(* Logix 5000 project; controller TFF vendor 1 type 14 code 107 rev 33.11; software revision 33.04; part 36 of 38 *)
(* tags used below, declared in another part *)
   Address : DINT;   // Temp Address
   AlarmInhibit_Timer : TIMER;
   Index : DINT;   // Index
   NewSystem : DINT;
   TIME : DINT[2];
   AI201B : ALIAS FOR AnalogPoint[0];
   AI201BAlarm : ALIAS FOR AlarmAnalog[0];
   AlarmAnalog_Storage : AlarmAnalog[6,50];
   AlarmDeviation : AlarmDeviation[20];   // Control Loop Deviation Alarm Array
   AlarmDeviation_Storage : AlarmDeviation[6,20];
   AnalogOutput_Storage : AnalogOutput[6,25];
   AnalogPoint_Storage : AnalogInput[6,50];
   CCPSystem : CCPSystem;   // CCP System Data
   CCPSystem_Storage : CCPSystem_Storage[6];
   ControlLoop : ControlLoop[20];   // Control Loop Array
   ControlLoop_Storage : ControlLoop[6,20];
   DigitalPoint_Storage : DigitalPoint[6,150];
   Drive : Drive[11];   // Drives Array
   Drive_Storage : Drive[6,11];
   FlowPath : FlowPath[64];   // Flow Path Array
   FlowPath_Storage : FlowPath[6,64];
   Gateway : Gateway;   // Gateway Control
   GWModbus : IO_Station;   // Status of Gateway Modbus
   Options : Options;   // Options List
   Phase0 : ALIAS FOR Phase[0];   // Phase 0
   Phase0_Totalizer_Feed : ALIAS FOR PhaseTotalizer[0];   // Phase 0 Total Feed
   PhaseTotalizer : PhaseTotalizer[18];   // Phase Totalizers Array
   PhaseTotalizer_Storage : PhaseTotalizer[6,18];
   PipeAnimation : PipeAnimation;   // HMI Pipe Animation Array
   PipeStatValueHMI : INT[224];   // Pipe Animation Value For HMI
   PISL601 : ALIAS FOR DigitalPoint[0];
   Rack_ACT350_WI101_200L : IO_Station;   // Status of ACT350 200L
   Rack_ACT350_WI101_500L : IO_Station;   // Status of ACT350 500L
   Rack_Murr_Node0_Smart : IO_Station;   // Status of Node 0 Smart
   Rack_Murr_Node1_TFF20 : IO_Station;   // Status of Node 1 TFF20
   Rack_Murr_Node1_TFF40 : IO_Station;   // Status of Node 1 TFF40
   Rack_Murr_Node1_TFF80 : IO_Station;   // Status of Node 1 TFF80
   SIC001 : ALIAS FOR Drive[1];
   SIC001_AO : ALIAS FOR AnalogOutput[0];
   SIC002 : ALIAS FOR Drive[2];
   ThisSystem : SystemType;
   Valve_Storage : Valve[6,100];
   WI101 : ALIAS FOR AnalogPoint[15];
   XV001 : ALIAS FOR Valve[0];
(* Process, continued *)

ROUTINE PipeAnimationHMI   (* ladder *)
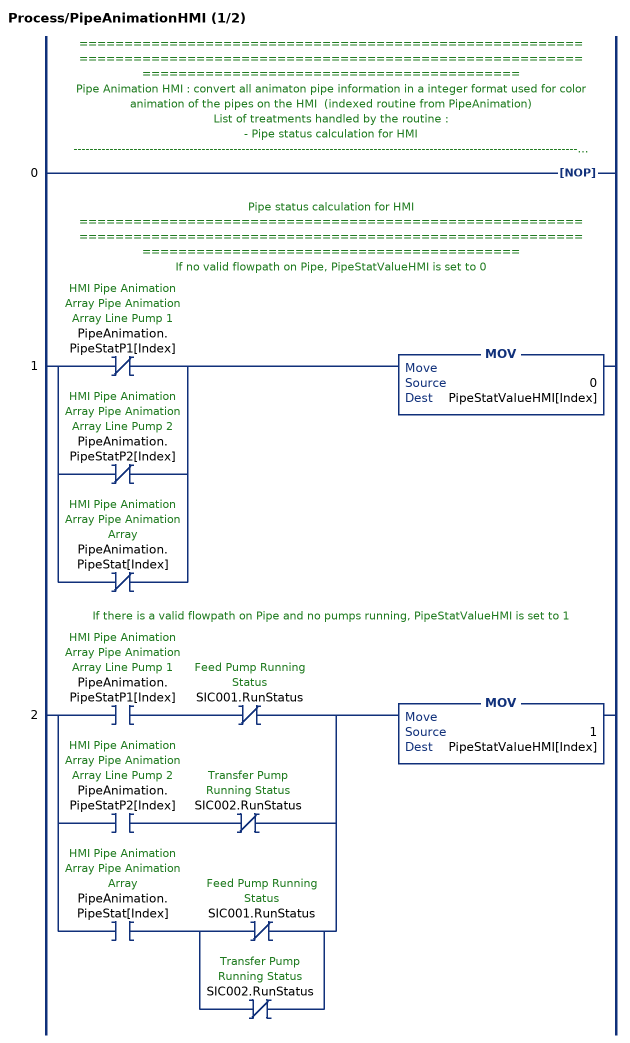
   // ==========================================================================================================================================================
   //                          Pipe Animation HMI : convert all animaton pipe information in a integer format used for color animation of the pipes on the HMI  (indexed routine from PipeAnimation)
   //                                                     List of treatments handled by the routine :
   //                                                          - Pipe status calculation for HMI
   //                                                     -----------------------------------------------------------------------------------------------------------------------------------------------------
   //                                                     History
   // 		2019-DEC-24 - Merck - Q. Spindler - Initial version for Candidate Release 1.00.00.00.a
   // ========================================================================================================================================================
   0: NOP();
   // Pipe status calculation for HMI
   // ==========================================================================================================================================================
   // If no valid flowpath on Pipe, PipeStatValueHMI is set to 0
   1: [XIO(PipeAnimation.PipeStatP1[Index]) ,XIO(PipeAnimation.PipeStatP2[Index]) ,XIO(PipeAnimation.PipeStat[Index]) ]MOV(0,PipeStatValueHMI[Index]);
   // If there is a valid flowpath on Pipe and no pumps running, PipeStatValueHMI is set to 1
   2: [XIC(PipeAnimation.PipeStatP1[Index]) XIO(SIC001.RunStatus) ,XIC(PipeAnimation.PipeStatP2[Index]) XIO(SIC002.RunStatus) ,XIC(PipeAnimation.PipeStat[Index]) [XIO(SIC001.RunStatus) ,XIO(SIC002.RunStatus) ] ]MOV(1,PipeStatValueHMI[Index]);
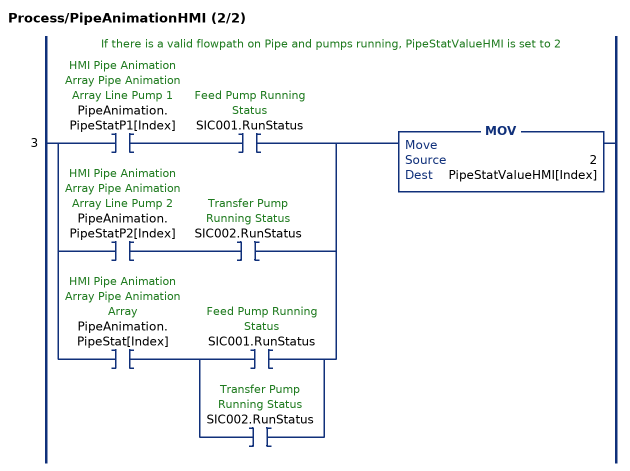
   // If there is a valid flowpath on Pipe and pumps running, PipeStatValueHMI is set to 2
   3: [XIC(PipeAnimation.PipeStatP1[Index]) XIC(SIC001.RunStatus) ,XIC(PipeAnimation.PipeStatP2[Index]) XIC(SIC002.RunStatus) ,XIC(PipeAnimation.PipeStat[Index]) [XIC(SIC001.RunStatus) ,XIC(SIC002.RunStatus) ] ]MOV(2,PipeStatValueHMI[Index]);
END_ROUTINE

ROUTINE Scale   (* function block diagram *)
// Scale Routine
   SHEET 1
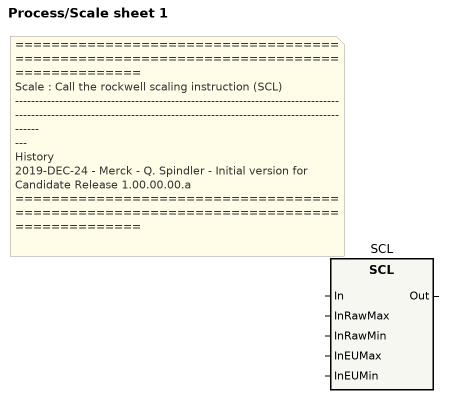
   // ======================================================================================
   // Scale : Call the rockwell scaling instruction (SCL)
   // ------------------------------------------------------------------------------------------------------------------------------------------------------------------------
   // ---
   // History
   // 	2019-DEC-24 - Merck - Q. Spindler - Initial version for Candidate Release 1.00.00.00.a
   // ======================================================================================
   SCL : SCL();   // unwired pins: In InRawMax InRawMin InEUMax InEUMin Out
END_ROUTINE

ROUTINE Station_Status   (* ladder *)
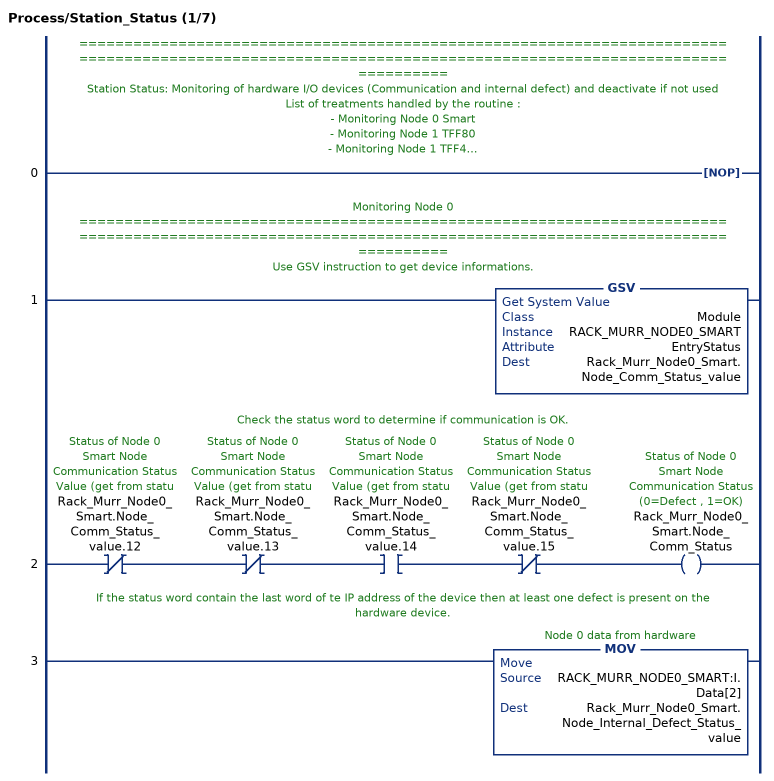
   // ==========================================================================================================================================================
   //                                                                   Station Status: Monitoring of hardware I/O devices (Communication and internal defect) and deactivate if not used
   //                                                     List of treatments handled by the routine :
   //                                                        - Monitoring Node 0 Smart
   //                                                        - Monitoring Node 1 TFF80
   //                                                        - Monitoring Node 1 TFF40
   //                                                        - Monitoring Node 1 TFF20
   //                                                       - Monitoring Modbus Gateway
   //                                                      - Monitoring ACT350 WI101 200L
   //                                                      - Monitoring ACT350 WI101 500L
   //                                                        - Deactivate / Activate devices
   //                                                     -----------------------------------------------------------------------------------------------------------------------------------------------------
   //                                                     History
   // 		2019-DEC-24 - Merck - Q. Spindler - Initial version for Candidate Release 1.00.00.00.a
   // ========================================================================================================================================================
   0: NOP();
   // Monitoring Node 0
   // ==========================================================================================================================================================
   // Use GSV instruction to get device informations.
   1: GSV(Module,RACK_MURR_NODE0_SMART,EntryStatus,Rack_Murr_Node0_Smart.Node_Comm_Status_value);
   // Check the status word to determine if communication is OK.
   2: XIO(Rack_Murr_Node0_Smart.Node_Comm_Status_value.12)XIO(Rack_Murr_Node0_Smart.Node_Comm_Status_value.13)XIC(Rack_Murr_Node0_Smart.Node_Comm_Status_value.14)XIO(Rack_Murr_Node0_Smart.Node_Comm_Status_value.15)OTE(Rack_Murr_Node0_Smart.Node_Comm_Status);
   // If the status word contain the last word of te IP address of the device then at least one defect is present on the hardware device.
   3: MOV(RACK_MURR_NODE0_SMART:I.Data[2],Rack_Murr_Node0_Smart.Node_Internal_Defect_Status_value);
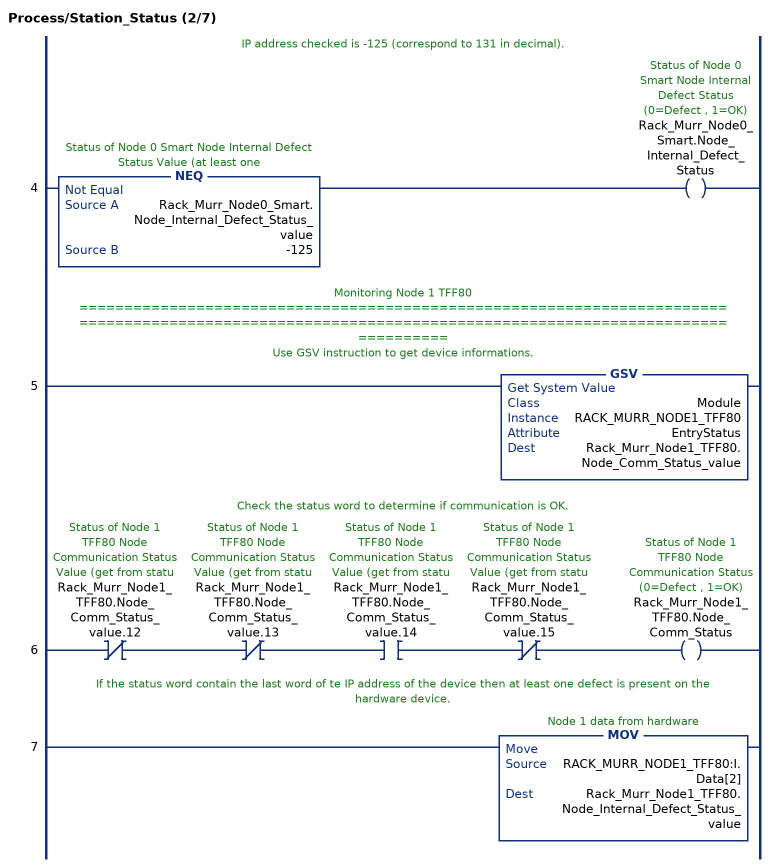
   // IP address checked is -125 (correspond to 131 in decimal).
   4: NEQ(Rack_Murr_Node0_Smart.Node_Internal_Defect_Status_value,-125)OTE(Rack_Murr_Node0_Smart.Node_Internal_Defect_Status);
   // Monitoring Node 1 TFF80
   // ==========================================================================================================================================================
   // Use GSV instruction to get device informations.
   5: GSV(Module,RACK_MURR_NODE1_TFF80,EntryStatus,Rack_Murr_Node1_TFF80.Node_Comm_Status_value);
   // Check the status word to determine if communication is OK.
   6: XIO(Rack_Murr_Node1_TFF80.Node_Comm_Status_value.12)XIO(Rack_Murr_Node1_TFF80.Node_Comm_Status_value.13)XIC(Rack_Murr_Node1_TFF80.Node_Comm_Status_value.14)XIO(Rack_Murr_Node1_TFF80.Node_Comm_Status_value.15)OTE(Rack_Murr_Node1_TFF80.Node_Comm_Status);
   // If the status word contain the last word of te IP address of the device then at least one defect is present on the hardware device.
   7: MOV(RACK_MURR_NODE1_TFF80:I.Data[2],Rack_Murr_Node1_TFF80.Node_Internal_Defect_Status_value);
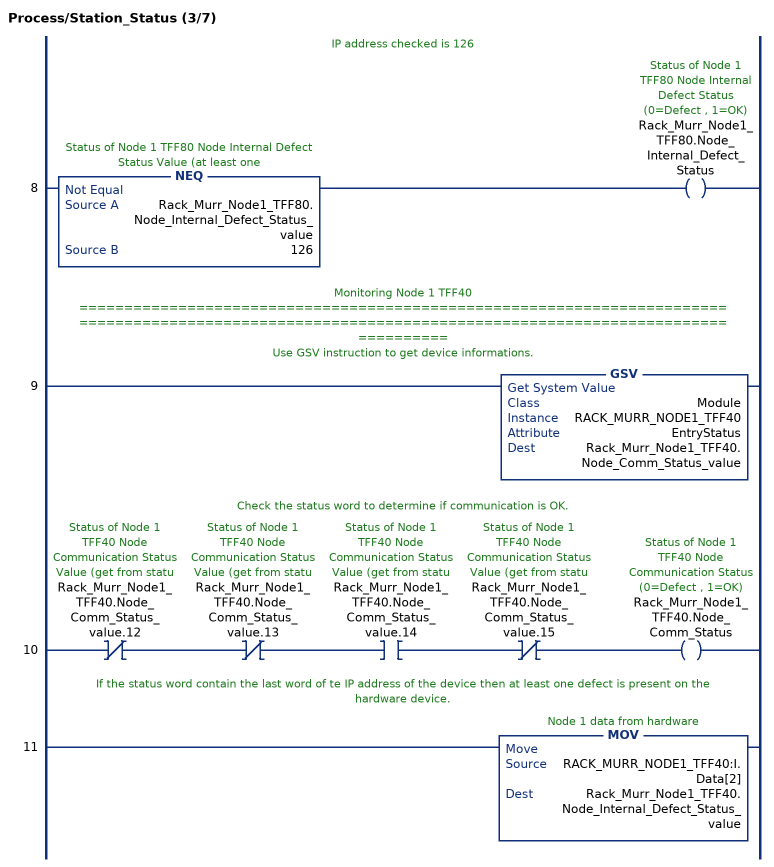
   // IP address checked is 126
   8: NEQ(Rack_Murr_Node1_TFF80.Node_Internal_Defect_Status_value,126)OTE(Rack_Murr_Node1_TFF80.Node_Internal_Defect_Status);
   // Monitoring Node 1 TFF40
   // ==========================================================================================================================================================
   // Use GSV instruction to get device informations.
   9: GSV(Module,RACK_MURR_NODE1_TFF40,EntryStatus,Rack_Murr_Node1_TFF40.Node_Comm_Status_value);
   // Check the status word to determine if communication is OK.
   10: XIO(Rack_Murr_Node1_TFF40.Node_Comm_Status_value.12)XIO(Rack_Murr_Node1_TFF40.Node_Comm_Status_value.13)XIC(Rack_Murr_Node1_TFF40.Node_Comm_Status_value.14)XIO(Rack_Murr_Node1_TFF40.Node_Comm_Status_value.15)OTE(Rack_Murr_Node1_TFF40.Node_Comm_Status);
   // If the status word contain the last word of te IP address of the device then at least one defect is present on the hardware device.
   11: MOV(RACK_MURR_NODE1_TFF40:I.Data[2],Rack_Murr_Node1_TFF40.Node_Internal_Defect_Status_value);
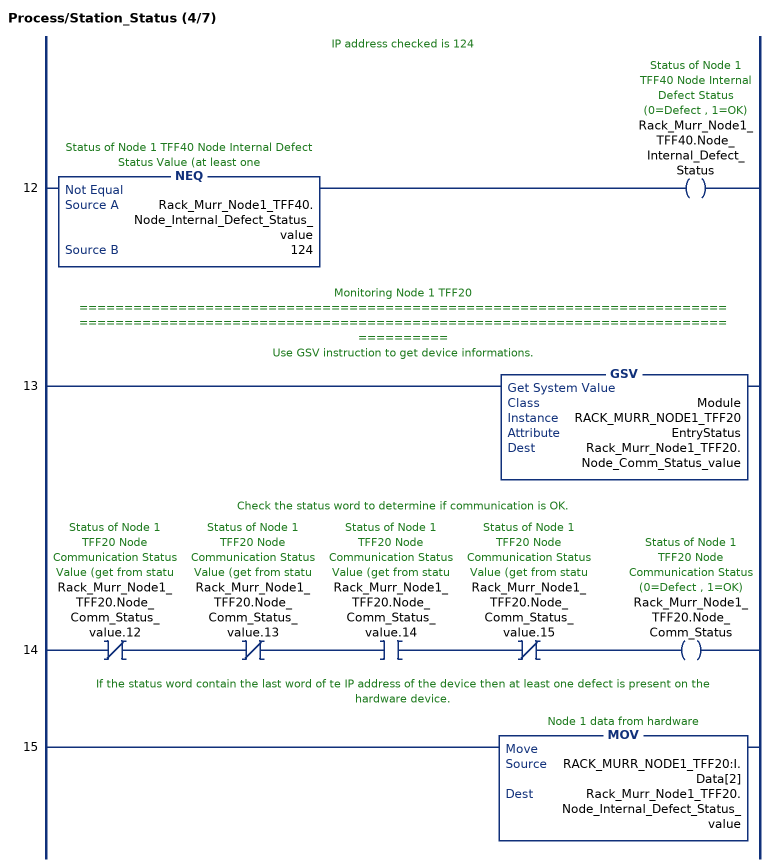
   // IP address checked is 124
   12: NEQ(Rack_Murr_Node1_TFF40.Node_Internal_Defect_Status_value,124)OTE(Rack_Murr_Node1_TFF40.Node_Internal_Defect_Status);
   // Monitoring Node 1 TFF20
   // ==========================================================================================================================================================
   // Use GSV instruction to get device informations.
   13: GSV(Module,RACK_MURR_NODE1_TFF20,EntryStatus,Rack_Murr_Node1_TFF20.Node_Comm_Status_value);
   // Check the status word to determine if communication is OK.
   14: XIO(Rack_Murr_Node1_TFF20.Node_Comm_Status_value.12)XIO(Rack_Murr_Node1_TFF20.Node_Comm_Status_value.13)XIC(Rack_Murr_Node1_TFF20.Node_Comm_Status_value.14)XIO(Rack_Murr_Node1_TFF20.Node_Comm_Status_value.15)OTE(Rack_Murr_Node1_TFF20.Node_Comm_Status);
   // If the status word contain the last word of te IP address of the device then at least one defect is present on the hardware device.
   15: MOV(RACK_MURR_NODE1_TFF20:I.Data[2],Rack_Murr_Node1_TFF20.Node_Internal_Defect_Status_value);
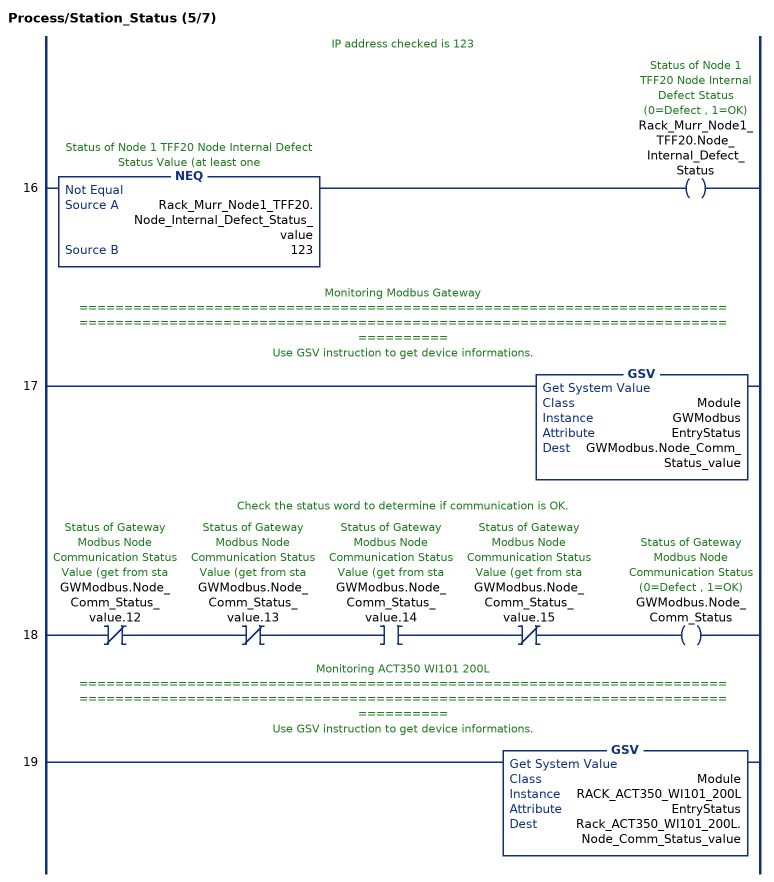
   // IP address checked is 123
   16: NEQ(Rack_Murr_Node1_TFF20.Node_Internal_Defect_Status_value,123)OTE(Rack_Murr_Node1_TFF20.Node_Internal_Defect_Status);
   // Monitoring Modbus Gateway
   // ==========================================================================================================================================================
   // Use GSV instruction to get device informations.
   17: GSV(Module,GWModbus,EntryStatus,GWModbus.Node_Comm_Status_value);
   // Check the status word to determine if communication is OK.
   18: XIO(GWModbus.Node_Comm_Status_value.12)XIO(GWModbus.Node_Comm_Status_value.13)XIC(GWModbus.Node_Comm_Status_value.14)XIO(GWModbus.Node_Comm_Status_value.15)OTE(GWModbus.Node_Comm_Status);
   // Monitoring ACT350 WI101 200L
   // ==========================================================================================================================================================
   // Use GSV instruction to get device informations.
   19: GSV(Module,RACK_ACT350_WI101_200L,EntryStatus,Rack_ACT350_WI101_200L.Node_Comm_Status_value);
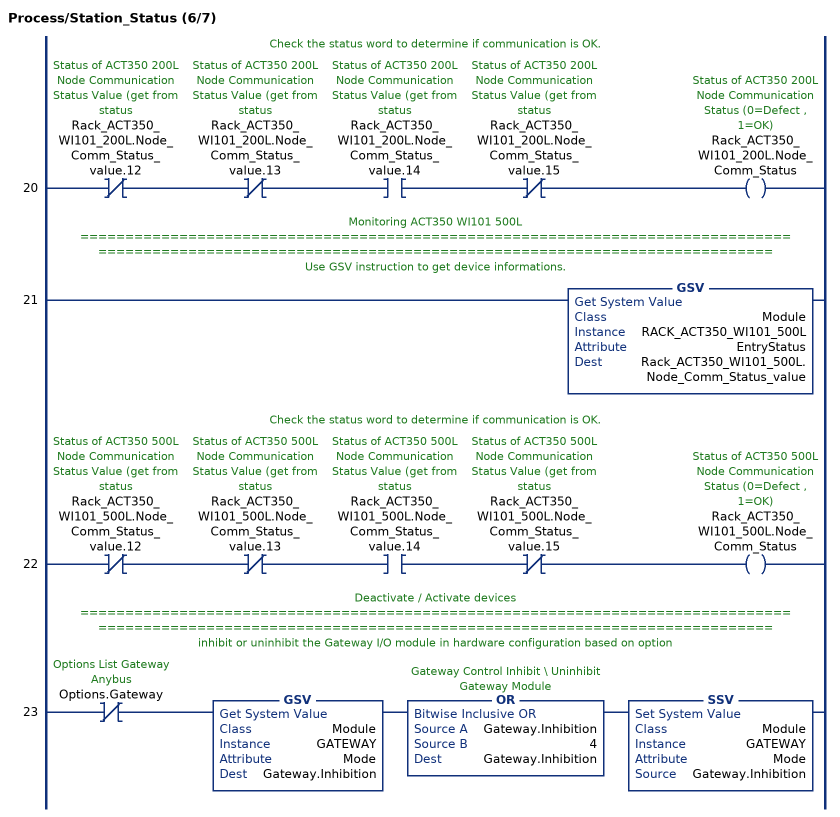
   // Check the status word to determine if communication is OK.
   20: XIO(Rack_ACT350_WI101_200L.Node_Comm_Status_value.12)XIO(Rack_ACT350_WI101_200L.Node_Comm_Status_value.13)XIC(Rack_ACT350_WI101_200L.Node_Comm_Status_value.14)XIO(Rack_ACT350_WI101_200L.Node_Comm_Status_value.15)OTE(Rack_ACT350_WI101_200L.Node_Comm_Status);
   // Monitoring ACT350 WI101 500L
   // ==========================================================================================================================================================
   // Use GSV instruction to get device informations.
   21: GSV(Module,RACK_ACT350_WI101_500L,EntryStatus,Rack_ACT350_WI101_500L.Node_Comm_Status_value);
   // Check the status word to determine if communication is OK.
   22: XIO(Rack_ACT350_WI101_500L.Node_Comm_Status_value.12)XIO(Rack_ACT350_WI101_500L.Node_Comm_Status_value.13)XIC(Rack_ACT350_WI101_500L.Node_Comm_Status_value.14)XIO(Rack_ACT350_WI101_500L.Node_Comm_Status_value.15)OTE(Rack_ACT350_WI101_500L.Node_Comm_Status);
   // Deactivate / Activate devices
   // ==========================================================================================================================================================
   // inhibit or uninhibit the Gateway I/O module in hardware configuration based on option
   23: XIO(Options.Gateway)GSV(Module,GATEWAY,Mode,Gateway.Inhibition)OR(Gateway.Inhibition,4,Gateway.Inhibition)SSV(Module,GATEWAY,Mode,Gateway.Inhibition);
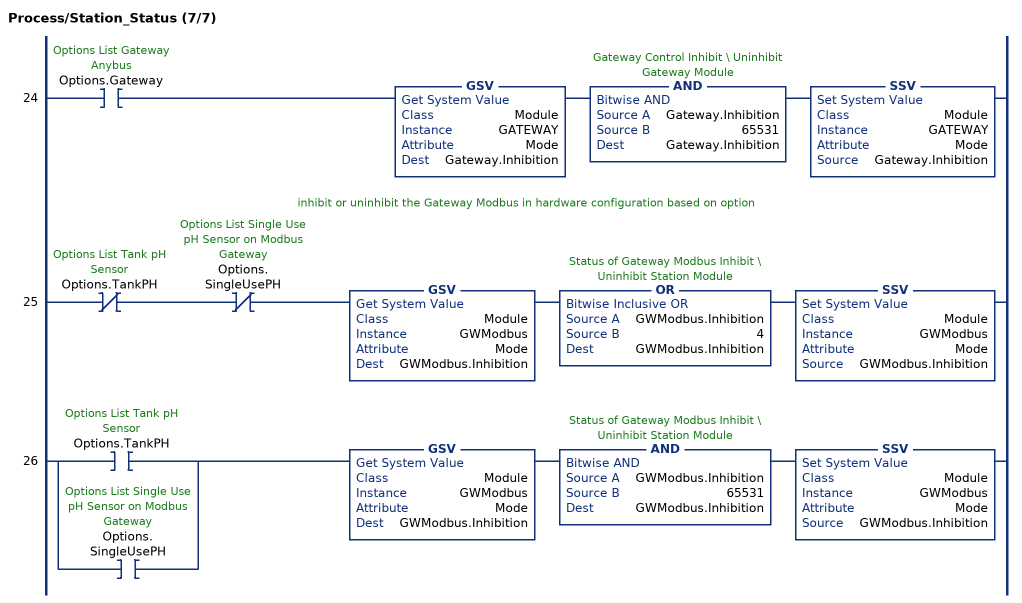
   24: XIC(Options.Gateway)GSV(Module,GATEWAY,Mode,Gateway.Inhibition)AND(Gateway.Inhibition,65531,Gateway.Inhibition)SSV(Module,GATEWAY,Mode,Gateway.Inhibition);
   // inhibit or uninhibit the Gateway Modbus in hardware configuration based on option
   25: XIO(Options.TankPH)XIO(Options.SingleUsePH)GSV(Module,GWModbus,Mode,GWModbus.Inhibition)OR(GWModbus.Inhibition,4,GWModbus.Inhibition)SSV(Module,GWModbus,Mode,GWModbus.Inhibition);
   26: [XIC(Options.TankPH) ,XIC(Options.SingleUsePH) ]GSV(Module,GWModbus,Mode,GWModbus.Inhibition)AND(GWModbus.Inhibition,65531,GWModbus.Inhibition)SSV(Module,GWModbus,Mode,GWModbus.Inhibition);
END_ROUTINE

ROUTINE SystemType   (* ladder *)
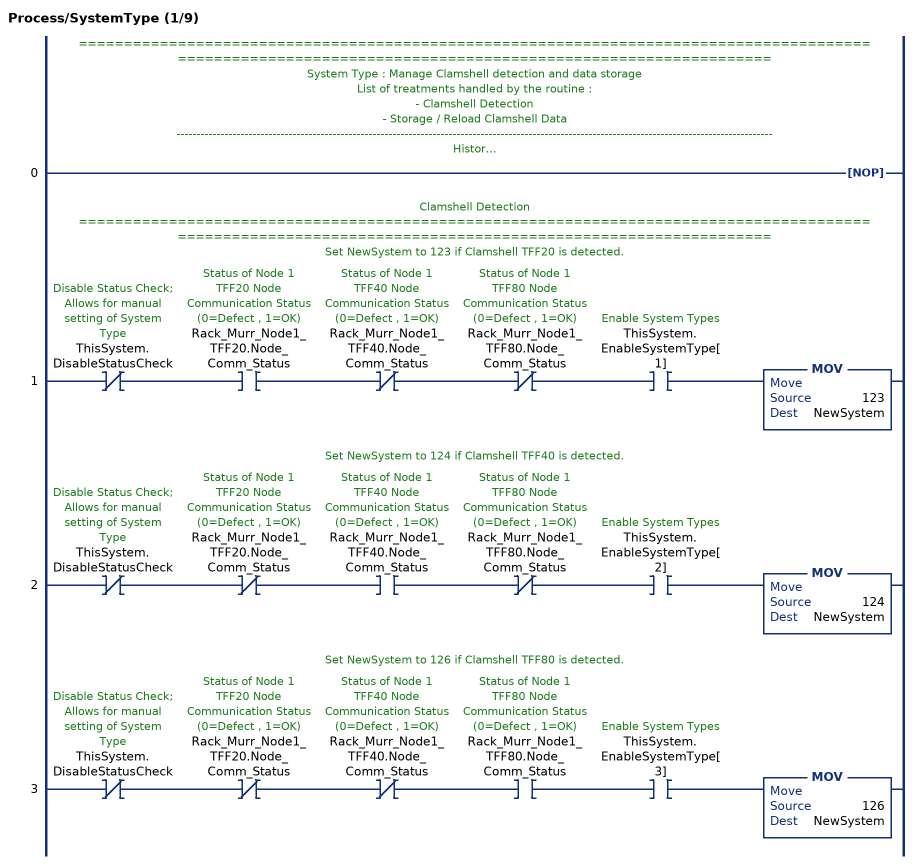
   // ==========================================================================================================================================================
   //                                                               System Type : Manage Clamshell detection and data storage
   //                                                     List of treatments handled by the routine :
   //                                                          - Clamshell Detection
   //                                                          - Storage / Reload Clamshell Data
   //                                                     -----------------------------------------------------------------------------------------------------------------------------------------------------
   //                                                     History
   // 		2019-DEC-24 - Merck - Q. Spindler - Initial version for Candidate Release 1.00.00.00.a
   //                                2022-JAN-11 - Merck - Q. Spindler - Modifications for Candidate Release 1.01.00.00.a
   // - Change PhaseTotalizer[0] lenght to 18
   // ========================================================================================================================================================
   0: NOP();
   // Clamshell Detection
   // ==========================================================================================================================================================
   // Set NewSystem to 123 if Clamshell TFF20 is detected.
   1: XIO(ThisSystem.DisableStatusCheck)XIC(Rack_Murr_Node1_TFF20.Node_Comm_Status)XIO(Rack_Murr_Node1_TFF40.Node_Comm_Status)XIO(Rack_Murr_Node1_TFF80.Node_Comm_Status)XIC(ThisSystem.EnableSystemType[1])MOV(123,NewSystem);
   // Set NewSystem to 124 if Clamshell TFF40 is detected.
   2: XIO(ThisSystem.DisableStatusCheck)XIO(Rack_Murr_Node1_TFF20.Node_Comm_Status)XIC(Rack_Murr_Node1_TFF40.Node_Comm_Status)XIO(Rack_Murr_Node1_TFF80.Node_Comm_Status)XIC(ThisSystem.EnableSystemType[2])MOV(124,NewSystem);
   // Set NewSystem to 126 if Clamshell TFF80 is detected.
   3: XIO(ThisSystem.DisableStatusCheck)XIO(Rack_Murr_Node1_TFF20.Node_Comm_Status)XIO(Rack_Murr_Node1_TFF40.Node_Comm_Status)XIC(Rack_Murr_Node1_TFF80.Node_Comm_Status)XIC(ThisSystem.EnableSystemType[3])MOV(126,NewSystem);
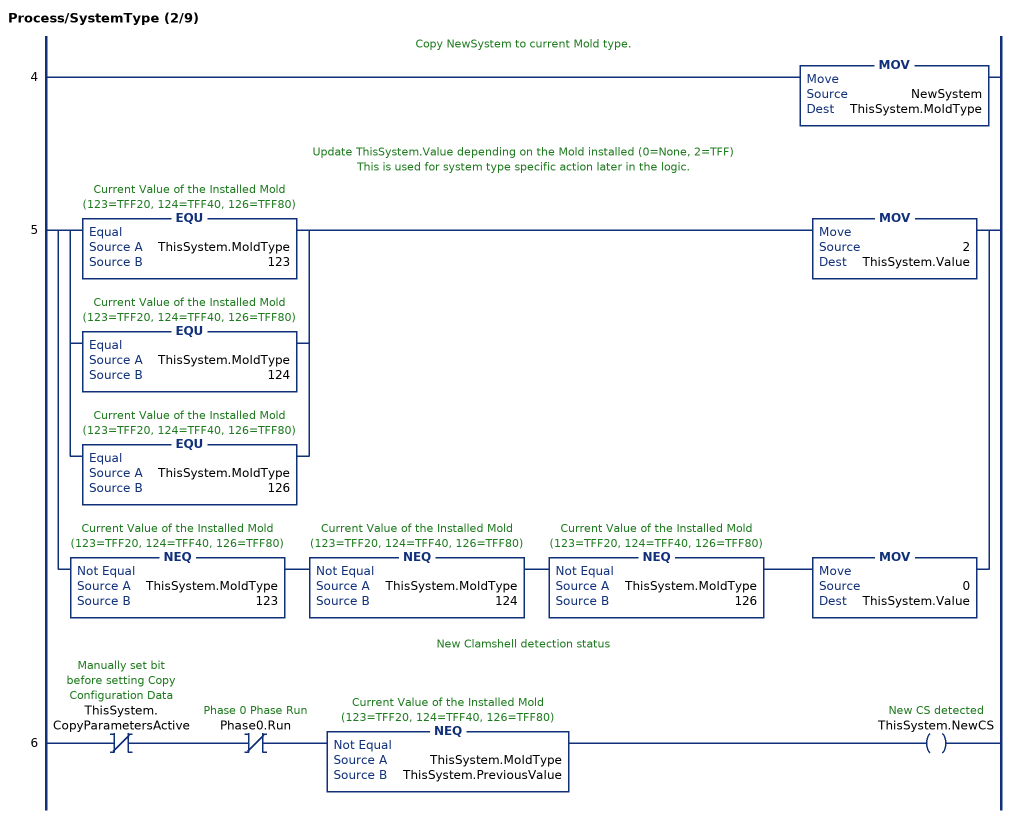
   // Copy NewSystem to current Mold type.
   4: MOV(NewSystem,ThisSystem.MoldType);
   // Update ThisSystem.Value depending on the Mold installed (0=None, 2=TFF)
   // This is used for system type specific action later in the logic.
   5: [[EQU(ThisSystem.MoldType,123) ,EQU(ThisSystem.MoldType,124) ,EQU(ThisSystem.MoldType,126) ] MOV(2,ThisSystem.Value) ,NEQ(ThisSystem.MoldType,123) NEQ(ThisSystem.MoldType,124) NEQ(ThisSystem.MoldType,126) MOV(0,ThisSystem.Value) ];
   // New Clamshell detection status
   6: XIO(ThisSystem.CopyParametersActive)XIO(Phase0.Run)NEQ(ThisSystem.MoldType,ThisSystem.PreviousValue)OTE(ThisSystem.NewCS);
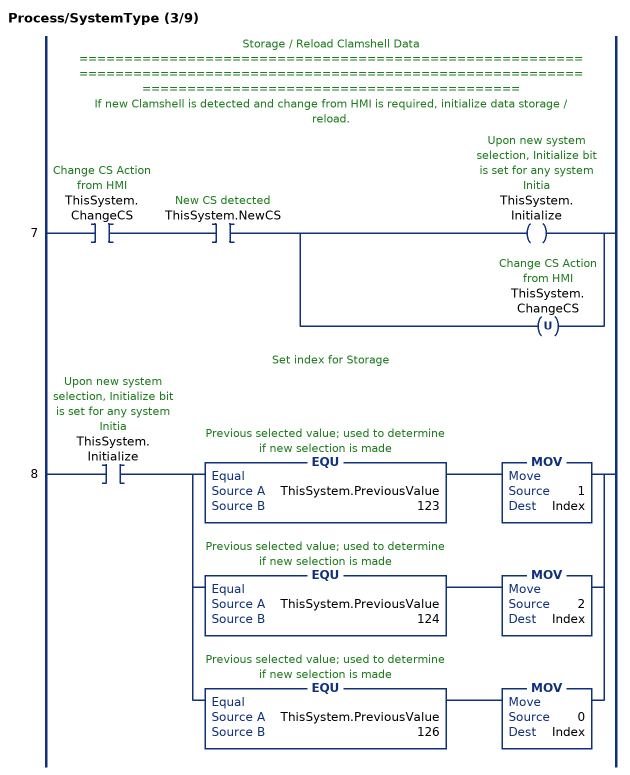
   // Storage / Reload Clamshell Data
   // ==========================================================================================================================================================
   // If new Clamshell is detected and change from HMI is required, initialize data storage / reload.
   7: XIC(ThisSystem.ChangeCS)XIC(ThisSystem.NewCS)[OTE(ThisSystem.Initialize) ,OTU(ThisSystem.ChangeCS) ];
   // Set index for Storage
   8: XIC(ThisSystem.Initialize)[EQU(ThisSystem.PreviousValue,123) MOV(1,Index) ,EQU(ThisSystem.PreviousValue,124) MOV(2,Index) ,EQU(ThisSystem.PreviousValue,126) MOV(0,Index) ];
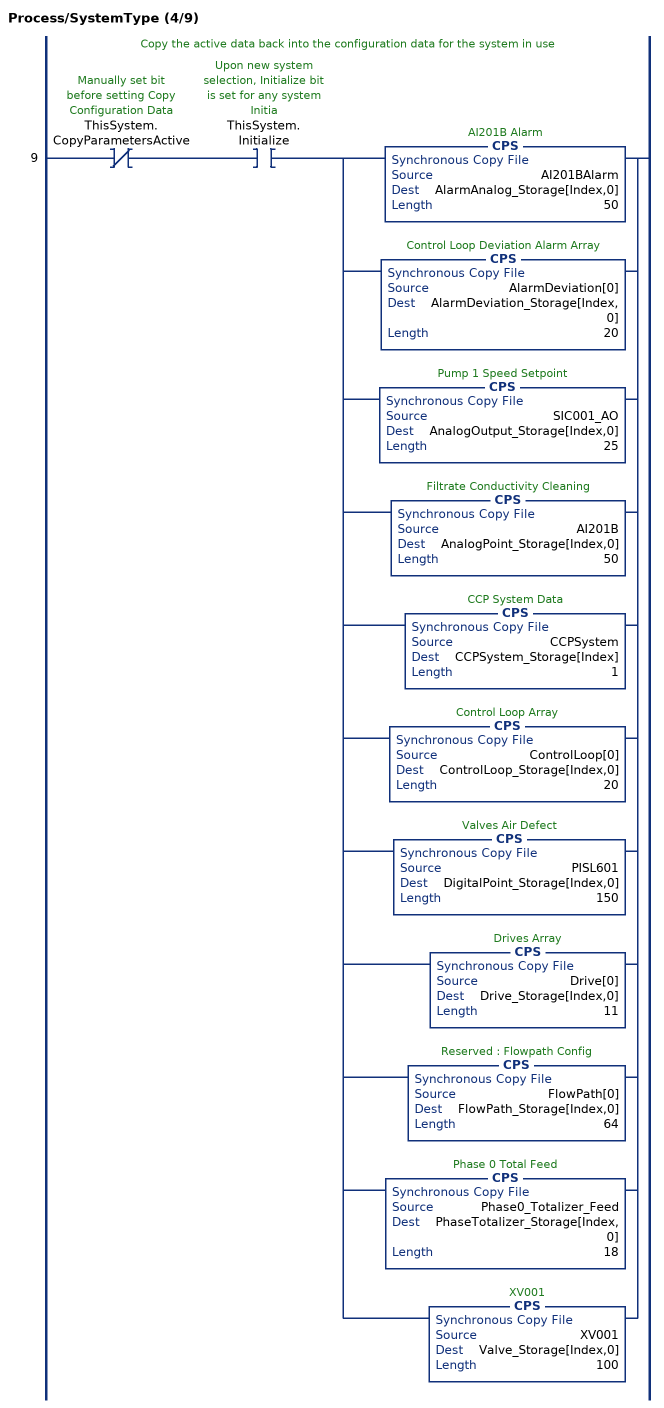
   // Copy the active data back into the configuration data for the system in use
   9: XIO(ThisSystem.CopyParametersActive)XIC(ThisSystem.Initialize)[CPS(AI201BAlarm,AlarmAnalog_Storage[Index,0],50) ,CPS(AlarmDeviation[0],AlarmDeviation_Storage[Index,0],20) ,CPS(SIC001_AO,AnalogOutput_Storage[Index,0],25) ,CPS(AI201B,AnalogPoint_Storage[Index,0],50) ,CPS(CCPSystem,CCPSystem_Storage[Index],1) ,CPS(ControlLoop[0],ControlLoop_Storage[Index,0],20) ,CPS(PISL601,DigitalPoint_Storage[Index,0],150) ,CPS(Drive[0],Drive_Storage[Index,0],11) ,CPS(FlowPath[0],FlowPath_Storage[Index,0],64) ,CPS(Phase0_Totalizer_Feed,PhaseTotalizer_Storage[Index,0],18) ,CPS(XV001,Valve_Storage[Index,0],100) ];
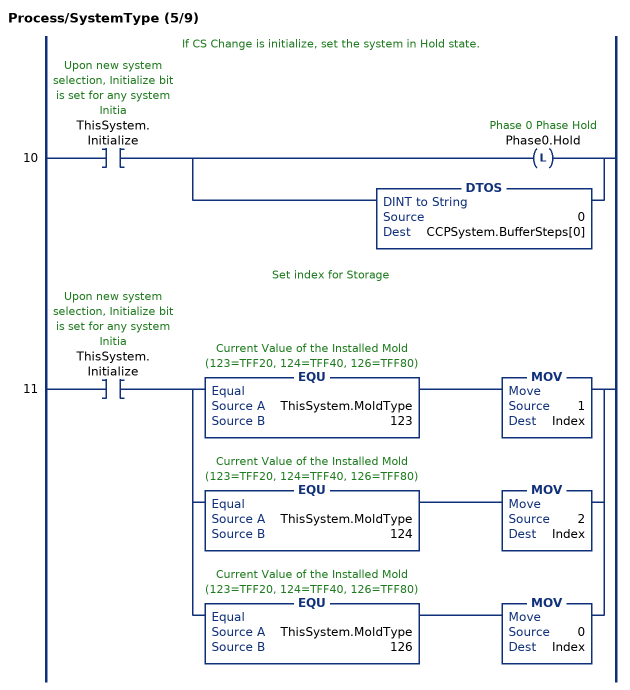
   // If CS Change is initialize, set the system in Hold state.
   10: XIC(ThisSystem.Initialize)[OTL(Phase0.Hold) ,DTOS(0,CCPSystem.BufferSteps[0]) ];
   // Set index for Storage
   11: XIC(ThisSystem.Initialize)[EQU(ThisSystem.MoldType,123) MOV(1,Index) ,EQU(ThisSystem.MoldType,124) MOV(2,Index) ,EQU(ThisSystem.MoldType,126) MOV(0,Index) ];
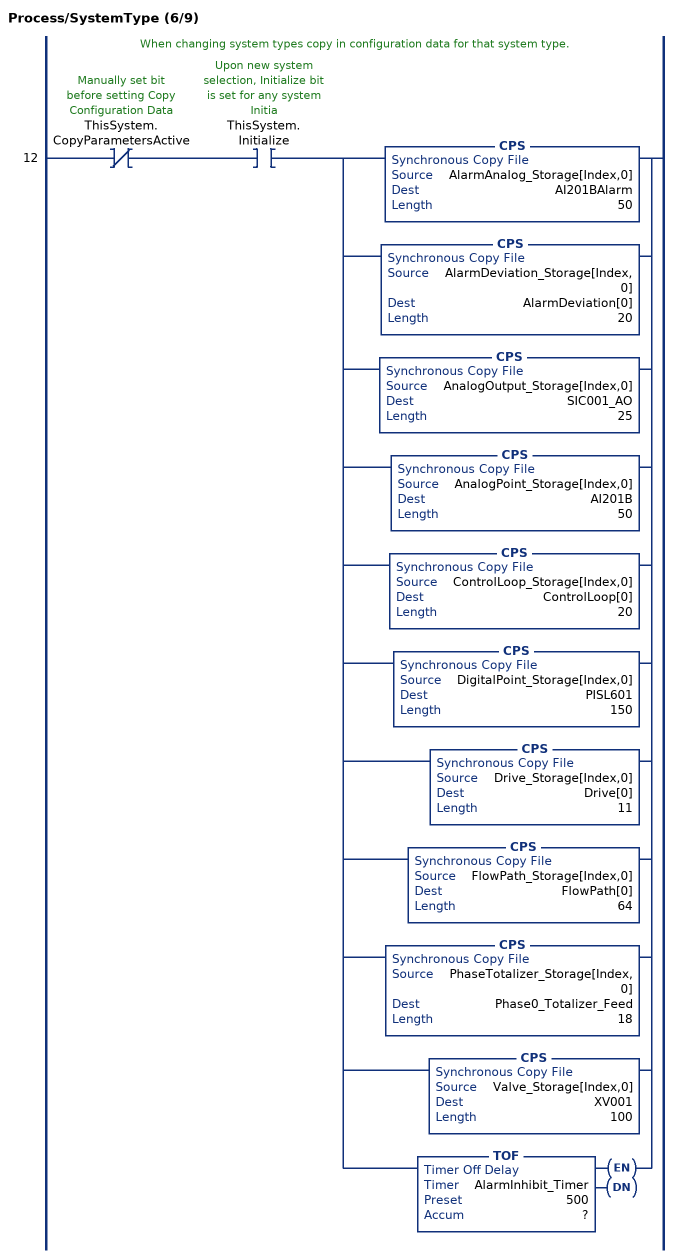
   // When changing system types copy in configuration data for that system type.
   12: XIO(ThisSystem.CopyParametersActive)XIC(ThisSystem.Initialize)[CPS(AlarmAnalog_Storage[Index,0],AI201BAlarm,50) ,CPS(AlarmDeviation_Storage[Index,0],AlarmDeviation[0],20) ,CPS(AnalogOutput_Storage[Index,0],SIC001_AO,25) ,CPS(AnalogPoint_Storage[Index,0],AI201B,50) ,CPS(ControlLoop_Storage[Index,0],ControlLoop[0],20) ,CPS(DigitalPoint_Storage[Index,0],PISL601,150) ,CPS(Drive_Storage[Index,0],Drive[0],11) ,CPS(FlowPath_Storage[Index,0],FlowPath[0],64) ,CPS(PhaseTotalizer_Storage[Index,0],Phase0_Totalizer_Feed,18) ,CPS(Valve_Storage[Index,0],XV001,100) ,TOF(AlarmInhibit_Timer,?,?) ];
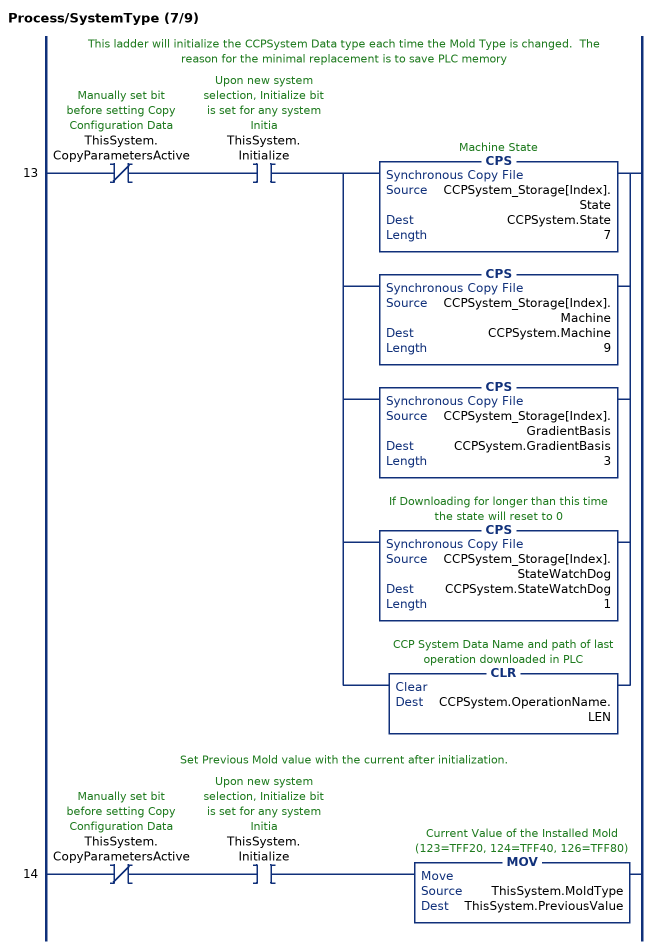
   // This ladder will initialize the CCPSystem Data type each time the Mold Type is changed.  The reason for the minimal replacement is to save PLC memory
   13: XIO(ThisSystem.CopyParametersActive)XIC(ThisSystem.Initialize)[CPS(CCPSystem_Storage[Index].State,CCPSystem.State,7) ,CPS(CCPSystem_Storage[Index].Machine,CCPSystem.Machine,9) ,CPS(CCPSystem_Storage[Index].GradientBasis,CCPSystem.GradientBasis,3) ,CPS(CCPSystem_Storage[Index].StateWatchDog,CCPSystem.StateWatchDog,1) ,CLR(CCPSystem.OperationName.LEN) ];
   // Set Previous Mold value with the current after initialization.
   14: XIO(ThisSystem.CopyParametersActive)XIC(ThisSystem.Initialize)MOV(ThisSystem.MoldType,ThisSystem.PreviousValue);
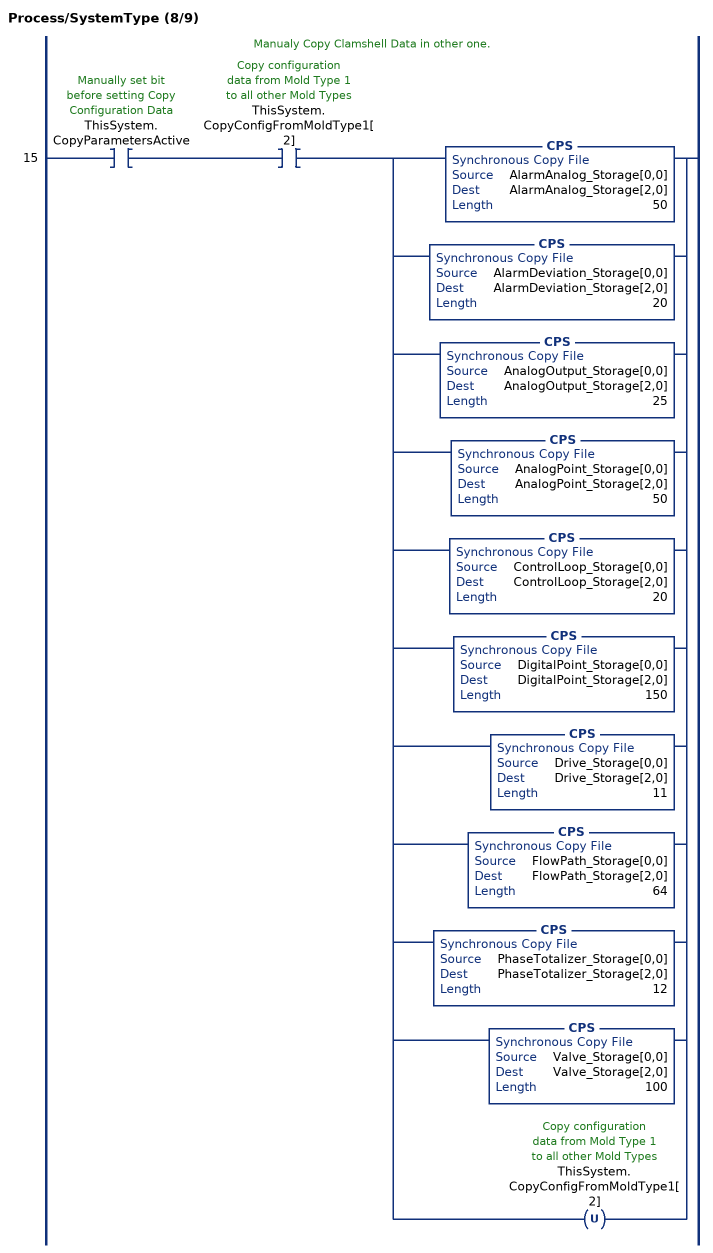
   // Manualy Copy Clamshell Data in other one.
   15: XIC(ThisSystem.CopyParametersActive)XIC(ThisSystem.CopyConfigFromMoldType1[2])[CPS(AlarmAnalog_Storage[0,0],AlarmAnalog_Storage[2,0],50) ,CPS(AlarmDeviation_Storage[0,0],AlarmDeviation_Storage[2,0],20) ,CPS(AnalogOutput_Storage[0,0],AnalogOutput_Storage[2,0],25) ,CPS(AnalogPoint_Storage[0,0],AnalogPoint_Storage[2,0],50) ,CPS(ControlLoop_Storage[0,0],ControlLoop_Storage[2,0],20) ,CPS(DigitalPoint_Storage[0,0],DigitalPoint_Storage[2,0],150) ,CPS(Drive_Storage[0,0],Drive_Storage[2,0],11) ,CPS(FlowPath_Storage[0,0],FlowPath_Storage[2,0],64) ,CPS(PhaseTotalizer_Storage[0,0],PhaseTotalizer_Storage[2,0],12) ,CPS(Valve_Storage[0,0],Valve_Storage[2,0],100) ,OTU(ThisSystem.CopyConfigFromMoldType1[2]) ];
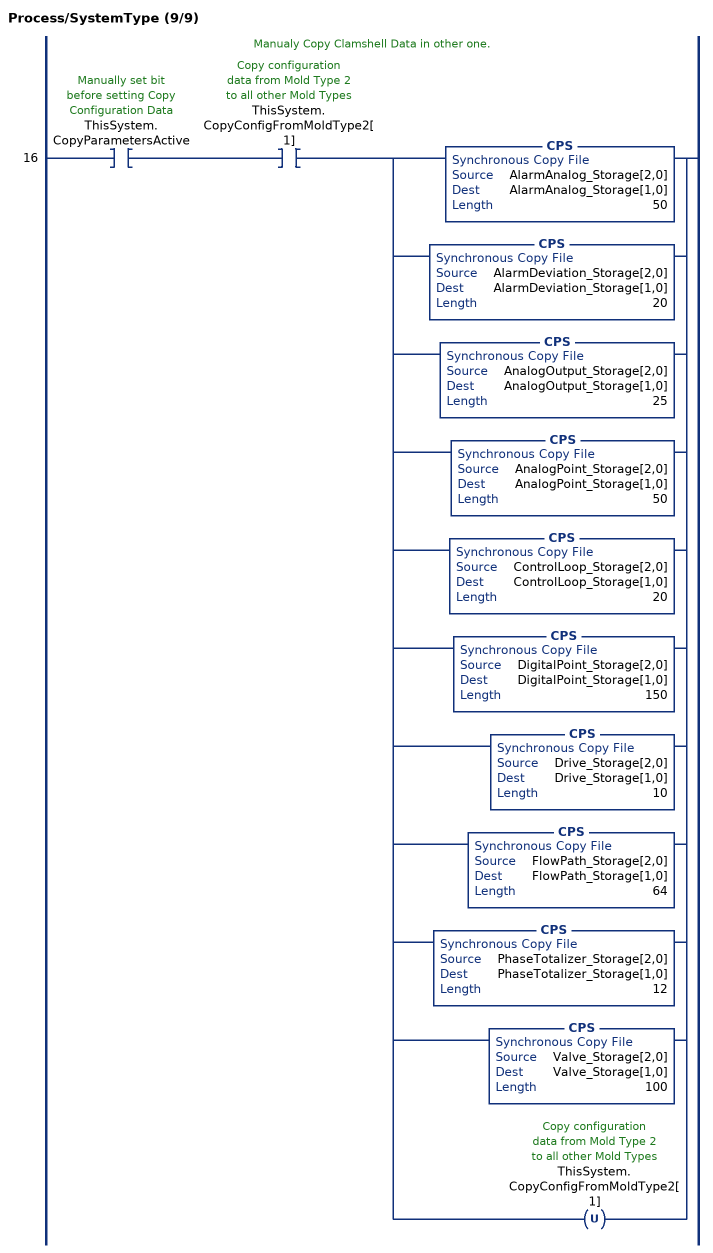
   // Manualy Copy Clamshell Data in other one.
   16: XIC(ThisSystem.CopyParametersActive)XIC(ThisSystem.CopyConfigFromMoldType2[1])[CPS(AlarmAnalog_Storage[2,0],AlarmAnalog_Storage[1,0],50) ,CPS(AlarmDeviation_Storage[2,0],AlarmDeviation_Storage[1,0],20) ,CPS(AnalogOutput_Storage[2,0],AnalogOutput_Storage[1,0],25) ,CPS(AnalogPoint_Storage[2,0],AnalogPoint_Storage[1,0],50) ,CPS(ControlLoop_Storage[2,0],ControlLoop_Storage[1,0],20) ,CPS(DigitalPoint_Storage[2,0],DigitalPoint_Storage[1,0],150) ,CPS(Drive_Storage[2,0],Drive_Storage[1,0],10) ,CPS(FlowPath_Storage[2,0],FlowPath_Storage[1,0],64) ,CPS(PhaseTotalizer_Storage[2,0],PhaseTotalizer_Storage[1,0],12) ,CPS(Valve_Storage[2,0],Valve_Storage[1,0],100) ,OTU(ThisSystem.CopyConfigFromMoldType2[1]) ];
END_ROUTINE
